(* PLC project Programme MGS_v0.3.10_Simulation.project, CODESYS CODESYS V3.5 SP19 Patch 1 *)
(* stored: creationDateTime 2026-07-04T07:57:21.9323215, modificationDateTime 2026-07-04T07:53:26.301727 *)

(* ═══════════════════════════════════════════════════════════════ ⚙️ ST_WinchHMI — Données d'échange IHM pour un treuil (M1/M2) ─────────────────────────────────────────────────────────────── 🎨 Destiné à l'affichage des bargraphes, LEDs, mesures et réglages. ═══════════════════════════════════════════════════════════════ *)
TYPE ST_WinchHMI : STRUCT
  TopSensorPositionM : REAL := 12.5;  (* 📐 Position cible du capteur haut (m) *)
  MaxStepDescente : INT := 2;  (* 🛑 Limitation palier vitesse en descente (1..5) *)
  RampAccelRate : REAL := 50;  (* 📈 Rampe d'accélération (%/s) *)
  RampDecelNormalRate : REAL := 150;  (* 📉 Rampe de décélération normale (%/s) *)
  RampDecelFastRate : REAL := 400;  (* ⚡ Rampe de décélération rapide / SafeStop (%/s) *)
  CableLimitDescentM : REAL := -20;  (* 📐 Limite basse physique de descente (m, négatif) *)
  SlowdownDistanceM : REAL := 1;  (* 📏 Distance avant limite pour enclencher le ralentissement (m) *)
  SlowSpeedPct : REAL := 15;  (* 📉 Vitesse de consigne lente dans la zone de ralentissement (%) *)
  PositionM : REAL;  (* 📊 Position actuelle du câble (mètres) *)
  SpeedRefPct : REAL;  (* 📈 Consigne de vitesse finale après rampe (%) *)
  StepNumber : INT;  (* 🔢 Palier de vitesse actif (0..5) *)
  FBState : E_State;  (* 🤖 État de l'automate interne (FB_Winch) *)
  Ready : BOOL;  (* 🟢 Treuil prêt à fonctionner *)
  Busy : BOOL;  (* ⚙️ Mouvement en cours *)
  Done : BOOL;  (* ✅ Action terminée *)
  Error : BOOL;  (* 🔴 Treuil en défaut *)
  ErrorId : WORD;  (* ❌ Code bitfield du défaut treuil *)
  RelayFwd : BOOL;  (* 🛗 Relais Montée activé *)
  RelayRev : BOOL;  (* 🛗 Relais Descente activé *)
  Contactor1 : BOOL;  (* 🔌 Contacteur vitesse palier 1 *)
  Contactor2 : BOOL;  (* 🔌 Contacteur vitesse palier 2 *)
  Contactor3 : BOOL;  (* 🔌 Contacteur vitesse palier 3 *)
  Contactor4 : BOOL;  (* 🔌 Contacteur vitesse palier 4 *)
  BrakeCmd : BOOL;  (* 🔓 Commande frein (TRUE = desserré / libre) *)
  Homed : BOOL;  (* 🎯 Prise d'origine (Homing) validée *)
  SafeStopActive : BOOL;  (* 🟧 Arrêt rapide activé par la sécurité *)
  ForbidDescentActive : BOOL;  (* 🚯 Descente interdite (détecteur mou de câble / limites) *)
  ForbidAscentActive : BOOL;  (* 🚯 Montée interdite (fin de course haut) *)
  SlackCableDetected : BOOL;  (* ⚠️ Mou de câble physiquement détecté *)
  ThermalFault : BOOL;  (* 🔥 Défaut surchauffe thermique moteur *)
  EncoderFault : BOOL;  (* 🔌 Perte de liaison ou incohérence codeur *)
  CableLimitDescentReached : BOOL;  (* ⚠️ Longueur max de câble atteinte (limite basse physique) *)
  Encoder : ST_EncoderHMI;  (* 🧲 Données d'échange et diagnostic du codeur *)
  FwdContactorCheck : ST_ContactorCheck;  (* 🔌 Coherence contacteur montée *)
  RevContactorCheck : ST_ContactorCheck;  (* 🔌 Coherence contacteur descente *)
  BrakeContactorCheck : ST_ContactorCheck;  (* 🔌 Coherence retour frein *)
  CmdReset : BOOL;  (* 🔑 Acquittement défauts spécifique treuil *)
  CmdHome : BOOL;  (* 🎯 Lancement de la prise d'origine *)
  ConfirmCoherence : BOOL;  (* 🔓 Confirmation de cohérence au démarrage *)
  BypassContactorFeedback : BOOL;  (* 🔌 Bypass retours contacteurs (banc de test) *)
  BypassSlackCable : BOOL;  (* ⚠️ Bypass capteur mou de câble (banc de test) *)
  BypassTopPositionSensor : BOOL;  (* 📐 Bypass capteur position haute (banc de test) *)
END_STRUCT;
END_TYPE
